(* IEC 61131-3 sources: Test-Git_ESME26/TestProgettoESME_26.fbsproj/AxisModuleLib Migration/AXM_FB_AxisModule.pou.xml.v3^ (part 2) *)

(* ---- Init_active.act.st ---- *)
__METADATA__
{
  "v3Meta": {
    "objectGuid": "f6f9ed11-c115-4c50-b3a9-4322940e64ce",
    "objectTypeGuid": "8ac092e5-3128-4e26-9e7e-11016c6684f2",
    "embeddedObjectTypeGuids": [
      "3b83b776-fb25-43b8-99f2-3c507c9143fc"
    ],
    "properties": {},
    "subObjects": {}
  }
}

iq_stStandardModuleItf.q_xActive := FALSE;
iq_stStandardModuleItf.q_xReady := FALSE;
iq_stStandardModuleItf.q_etDiag := GD.ET_Diag.Ok;
iq_stStandardModuleItf.q_udiDiagExt := AXM_ET_DiagExt.Disabled;
iq_stStandardModuleItf.q_sDiagExt := AXM_FC_EtDiagExtToString(i_etDiagExt := iq_stStandardModuleItf.q_udiDiagExt);
iq_stStandardModuleItf.q_sMsg := AXM_FC_EtDiagExtToString(i_etDiagExt := AXM_ET_DiagExt.Disabled);
iq_stStandardModuleItf.q_dwModuleType := TPL.ET_ModuleType.AxisModule;
iq_stStandardModuleItf.q_sModuleTypeName := 'AxisModule';
iq_stStandardModuleItf.q_udiModuleVersion := 1;

iq_stAxisModuleItf.stMain.q_etOpMode := AXM_ET_OpMode.NoOp;
iq_stAxisModuleItf.stMain.q_etState := AXM_ET_State.Disabled;

THIS^.DiagQuit();
THIS^.InactiveCMDExecution();

(* detect invalid configurations and avoid array index out of range error *)
IF(iq_stStandardModuleItf.iq_stExt.udiReactionOffset + TPL.ET_Reaction.MainsContactorOff > TPL.Gc_udiMaxNumberOfReactions) OR xExceptionReactionOutsideRange THEN (* module uses error reactions 1 to 5 *)
	xExceptionReactionOutsideRange := TRUE; (* create unquittable error *)
	(* create exception *)
	stExceptionInit.etDiag					:= GD.ET_Diag.InputParameterInvalid;
	stExceptionInit.udiDiagExt				:= AXM_ET_DiagExt.ReactionOffsetRange;
	stExceptionInit.sMsg					:= Standard.CONCAT('Value: ', UDINT_TO_STRING(iq_stStandardModuleItf.iq_stExt.udiReactionOffset));
	stExceptionInit.udiModuleId				:= iq_stStandardModuleItf.i_udiModuleId;
	stExceptionInit.sModuleName				:= iq_stStandardModuleItf.i_sModuleName;
	stExceptionInit.etSource				:= TPL.ET_ExceptionSource.AxisModule;
	stExceptionInit.timDelayTime			:= T#0MS;
	stExceptionInit.wHmiAttributes			:= 0;
	stExceptionInit.xAutoQuit				:= FALSE;
	stExceptionInit.stReaction.axReaction[TPL.ET_Reaction.AsyncStop]	:= TRUE; (* without offset on purpose *)
	iq_stStandardModuleItf.iq_stExt.udiReactionOffset := 0;
	ReportException(iq_stException := stExceptionInit);
ELSIF(iq_stStandardModuleItf.i_xEnable) THEN
	stReaction1 := stEmptyReaction;
	stReaction1.axReaction[iq_stStandardModuleItf.iq_stExt.udiReactionOffset + TPL.ET_Reaction.AsyncStop] := TRUE;
	stReaction2 := stEmptyReaction;
	stReaction2.axReaction[iq_stStandardModuleItf.iq_stExt.udiReactionOffset + TPL.ET_Reaction.SyncStopEL] := TRUE;
	stReaction3 := stEmptyReaction;
	stReaction3.axReaction[iq_stStandardModuleItf.iq_stExt.udiReactionOffset + TPL.ET_Reaction.SyncStopEH] := TRUE;
	stReaction4 := stEmptyReaction;
	stReaction4.axReaction[iq_stStandardModuleItf.iq_stExt.udiReactionOffset + TPL.ET_Reaction.StopEndOfCycle] := TRUE;

	(* Initialization of exception structures *)
	stExceptionCmdUnknown.etDiag			:= GD.ET_Diag.ExecutionAborted;
	stExceptionCmdUnknown.udiDiagExt		:= AXM_ET_DiagExt.CmdUnknown;
	stExceptionCmdUnknown.sMsg				:= 'Command unknown'; (* Replaced on usage *)
	stExceptionCmdUnknown.udiModuleId		:= iq_stStandardModuleItf.i_udiModuleId;
	stExceptionCmdUnknown.sModuleName		:= iq_stStandardModuleItf.i_sModuleName;
	stExceptionCmdUnknown.etSource			:= TPL.ET_ExceptionSource.AxisModule;
	stExceptionCmdUnknown.timDelayTime		:= T#0MS;
	stExceptionCmdUnknown.wHmiAttributes	:= 0;
	stExceptionCmdUnknown.xAutoQuit			:= FALSE;
	stExceptionCmdUnknown.stReaction		:= stReaction1;

	stExceptionCmdImpossibleOverwrite.etDiag			:= GD.ET_Diag.ExecutionAborted;
	stExceptionCmdImpossibleOverwrite.udiDiagExt		:= AXM_ET_DiagExt.CmdImpossibleOverwrite;
	stExceptionCmdImpossibleOverwrite.sMsg				:= 'Impossible command overwrite'; (* Replaced on usage *)
	stExceptionCmdImpossibleOverwrite.udiModuleId		:= iq_stStandardModuleItf.i_udiModuleId;
	stExceptionCmdImpossibleOverwrite.sModuleName		:= iq_stStandardModuleItf.i_sModuleName;
	stExceptionCmdImpossibleOverwrite.etSource			:= TPL.ET_ExceptionSource.AxisModule;
	stExceptionCmdImpossibleOverwrite.timDelayTime		:= T#0MS;
	stExceptionCmdImpossibleOverwrite.wHmiAttributes	:= 0;
	stExceptionCmdImpossibleOverwrite.xAutoQuit			:= FALSE;
	stExceptionCmdImpossibleOverwrite.stReaction		:= stReaction1;

	stExceptionCmdImpossibleState.etDiag			:= GD.ET_Diag.ExecutionAborted;
	stExceptionCmdImpossibleState.udiDiagExt		:= AXM_ET_DiagExt.CmdImpossibleState;
	stExceptionCmdImpossibleState.sMsg				:= 'Impossible command for state'; (* Replaced on usage *)
	stExceptionCmdImpossibleState.udiModuleId		:= iq_stStandardModuleItf.i_udiModuleId;
	stExceptionCmdImpossibleState.sModuleName		:= iq_stStandardModuleItf.i_sModuleName;
	stExceptionCmdImpossibleState.etSource			:= TPL.ET_ExceptionSource.AxisModule;
	stExceptionCmdImpossibleState.timDelayTime		:= T#0MS;
	stExceptionCmdImpossibleState.wHmiAttributes	:= 0;
	stExceptionCmdImpossibleState.xAutoQuit			:= FALSE;
	stExceptionCmdImpossibleState.stReaction		:= stReaction1;

	stWarningCmdImpossibleReaction.etDiag			:= GD.ET_Diag.ExecutionAborted;
	stWarningCmdImpossibleReaction.udiDiagExt		:= AXM_ET_DiagExt.CmdImpossibleReaction;
	stWarningCmdImpossibleReaction.sMsg				:= 'Impossible command on reaction'; (* Replaced on usage *)
	stWarningCmdImpossibleReaction.udiModuleId		:= iq_stStandardModuleItf.i_udiModuleId;
	stWarningCmdImpossibleReaction.sModuleName		:= iq_stStandardModuleItf.i_sModuleName;
	stWarningCmdImpossibleReaction.etSource			:= TPL.ET_ExceptionSource.AxisModule;
	stWarningCmdImpossibleReaction.timDelayTime	:= T#0MS;
	stWarningCmdImpossibleReaction.wHmiAttributes	:= 0;
	stWarningCmdImpossibleReaction.xAutoQuit		:= FALSE;

	stExceptionDriveFatal.etDiag			:= GD.ET_Diag.DriveConditionInvalid;
	stExceptionDriveFatal.udiDiagExt		:= AXM_ET_DiagExt.DriveExceptionFatal;
	stExceptionDriveFatal.sMsg				:= 'Drive diag'; (* Replaced on usage *)
	stExceptionDriveFatal.udiModuleId		:= iq_stStandardModuleItf.i_udiModuleId;
	stExceptionDriveFatal.sModuleName		:= iq_stStandardModuleItf.i_sModuleName;
	stExceptionDriveFatal.etSource			:= TPL.ET_ExceptionSource.AxisModule;
	stExceptionDriveFatal.timDelayTime		:= T#0MS;
	stExceptionDriveFatal.wHmiAttributes	:= 0;
	stExceptionDriveFatal.xAutoQuit			:= FALSE;
	stExceptionDriveFatal.stReaction		:= stReaction1;

	stExcepitonDrive.etDiag			:= GD.ET_Diag.DriveConditionInvalid;
	stExcepitonDrive.udiDiagExt		:= AXM_ET_DiagExt.DriveException;
	stExcepitonDrive.sMsg			:= 'Drive diag'; (* Replaced on usage *)
	stExcepitonDrive.udiModuleId	:= iq_stStandardModuleItf.i_udiModuleId;
	stExcepitonDrive.sModuleName	:= iq_stStandardModuleItf.i_sModuleName;
	stExcepitonDrive.etSource		:= TPL.ET_ExceptionSource.AxisModule;
	stExcepitonDrive.timDelayTime	:= T#0MS;
	stExcepitonDrive.wHmiAttributes	:= 0;
	stExcepitonDrive.xAutoQuit		:= FALSE;
	stExcepitonDrive.stReaction		:= stReaction2;

	stWarningDrive.etDiag			:= GD.ET_Diag.DriveConditionInvalid;
	stWarningDrive.udiDiagExt		:= AXM_ET_DiagExt.DriveWarning;
	stWarningDrive.sMsg				:= 'Drive warning'; (* Replaced on usage *)
	stWarningDrive.udiModuleId		:= iq_stStandardModuleItf.i_udiModuleId;
	stWarningDrive.sModuleName		:= iq_stStandardModuleItf.i_sModuleName;
	stWarningDrive.etSource			:= TPL.ET_ExceptionSource.AxisModule;
	stWarningDrive.timDelayTime		:= T#0MS;
	stWarningDrive.wHmiAttributes	:= 0;
	stWarningDrive.xAutoQuit		:= FALSE;
	stWarningDrive.stReaction		:= stReaction4;

	stExceptionPosHwLimit.etDiag			:= GD.ET_Diag.LimitReached;
	stExceptionPosHwLimit.udiDiagExt		:= AXM_ET_DiagExt.HwLimitPosReached;
	stExceptionPosHwLimit.sMsg				:= '';
	stExceptionPosHwLimit.udiModuleId		:= iq_stStandardModuleItf.i_udiModuleId;
	stExceptionPosHwLimit.sModuleName		:= iq_stStandardModuleItf.i_sModuleName;
	stExceptionPosHwLimit.etSource			:= TPL.ET_ExceptionSource.AxisModule;
	stExceptionPosHwLimit.timDelayTime		:= T#0MS;
	stExceptionPosHwLimit.wHmiAttributes	:= 0;
	stExceptionPosHwLimit.xAutoQuit			:= FALSE;
	stExceptionPosHwLimit.stReaction		:= stReaction3;

	stExceptionNegHwLimit.etDiag			:= GD.ET_Diag.LimitReached;
	stExceptionNegHwLimit.udiDiagExt		:= AXM_ET_DiagExt.HwLimitNegReached;
	stExceptionNegHwLimit.sMsg				:= '';
	stExceptionNegHwLimit.udiModuleId		:= iq_stStandardModuleItf.i_udiModuleId;
	stExceptionNegHwLimit.sModuleName		:= iq_stStandardModuleItf.i_sModuleName;
	stExceptionNegHwLimit.etSource			:= TPL.ET_ExceptionSource.AxisModule;
	stExceptionNegHwLimit.timDelayTime		:= T#0MS;
	stExceptionNegHwLimit.wHmiAttributes	:= 0;
	stExceptionNegHwLimit.xAutoQuit			:= FALSE;
	stExceptionNegHwLimit.stReaction		:= stReaction3;

	stWarningPosHwLimit.etDiag			:= GD.ET_Diag.LimitReached;
	stWarningPosHwLimit.udiDiagExt		:= AXM_ET_DiagExt.HwLimitPosWarning;
	stWarningPosHwLimit.sMsg			:= '';
	stWarningPosHwLimit.udiModuleId		:= iq_stStandardModuleItf.i_udiModuleId;
	stWarningPosHwLimit.sModuleName		:= iq_stStandardModuleItf.i_sModuleName;
	stWarningPosHwLimit.etSource		:= TPL.ET_ExceptionSource.AxisModule;
	stWarningPosHwLimit.timDelayTime	:= T#0MS;
	stWarningPosHwLimit.wHmiAttributes	:= 0;
	stWarningPosHwLimit.xAutoQuit		:= TRUE;

	stWarningNegHwLimit.etDiag			:= GD.ET_Diag.LimitReached;
	stWarningNegHwLimit.udiDiagExt		:= AXM_ET_DiagExt.HwLimitNegWarning;
	stWarningNegHwLimit.sMsg			:= '';
	stWarningNegHwLimit.udiModuleId		:= iq_stStandardModuleItf.i_udiModuleId;
	stWarningNegHwLimit.sModuleName		:= iq_stStandardModuleItf.i_sModuleName;
	stWarningNegHwLimit.etSource		:= TPL.ET_ExceptionSource.AxisModule;
	stWarningNegHwLimit.timDelayTime	:= T#0MS;
	stWarningNegHwLimit.wHmiAttributes	:= 0;
	stWarningNegHwLimit.xAutoQuit		:= TRUE;

	stExceptionVelLimitCrossed.etDiag			:= GD.ET_Diag.LimitReached;
	stExceptionVelLimitCrossed.udiDiagExt		:= AXM_ET_DiagExt.ReducedVelocityLImit;
	stExceptionVelLimitCrossed.sMsg				:= '';
	stExceptionVelLimitCrossed.udiModuleId		:= iq_stStandardModuleItf.i_udiModuleId;
	stExceptionVelLimitCrossed.sModuleName		:= iq_stStandardModuleItf.i_sModuleName;
	stExceptionVelLimitCrossed.etSource			:= TPL.ET_ExceptionSource.AxisModule;
	stExceptionVelLimitCrossed.timDelayTime		:= T#0MS;
	stExceptionVelLimitCrossed.wHmiAttributes	:= 0;
	stExceptionVelLimitCrossed.xAutoQuit		:= FALSE;
	stExceptionVelLimitCrossed.stReaction		:= stReaction1;

	stExceptionUnexpected.etDiag			:= GD.ET_Diag.UnexpectedProgramBehavior;
	stExceptionUnexpected.udiDiagExt		:= AXM_ET_DiagExt.UnknownFeedback;
	stExceptionUnexpected.sMsg				:= ''; (* Replaced on usage *)
	stExceptionUnexpected.udiModuleId		:= iq_stStandardModuleItf.i_udiModuleId;
	stExceptionUnexpected.sModuleName		:= iq_stStandardModuleItf.i_sModuleName;
	stExceptionUnexpected.etSource			:= TPL.ET_ExceptionSource.AxisModule;
	stExceptionUnexpected.timDelayTime		:= T#0MS;
	stExceptionUnexpected.wHmiAttributes	:= 0;
	stExceptionUnexpected.xAutoQuit			:= FALSE;
	stExceptionUnexpected.stReaction		:= stReaction1;

	stExceptionModuleReaction1.etDiag			:= GD.ET_Diag.InputParameterInvalid;(* Replaced on usage *)
	stExceptionModuleReaction1.udiDiagExt		:= AXM_ET_DiagExt.DriveInvalid;(* Replaced on usage *)
	stExceptionModuleReaction1.sMsg				:= '';(* Replaced on usage *)
	stExceptionModuleReaction1.udiModuleId		:= iq_stStandardModuleItf.i_udiModuleId;
	stExceptionModuleReaction1.sModuleName		:= iq_stStandardModuleItf.i_sModuleName;
	stExceptionModuleReaction1.etSource			:= TPL.ET_ExceptionSource.AxisModule;
	stExceptionModuleReaction1.timDelayTime		:= T#0MS;
	stExceptionModuleReaction1.wHmiAttributes	:= 0;
	stExceptionModuleReaction1.xAutoQuit		:= FALSE;
	stExceptionModuleReaction1.stReaction		:= stReaction1;

	stExceptionModuleReaction2.etDiag			:= GD.ET_Diag.InputParameterInvalid;(* Replaced on usage *)
	stExceptionModuleReaction2.udiDiagExt		:= AXM_ET_DiagExt.DriveInvalid;(* Replaced on usage *)
	stExceptionModuleReaction2.sMsg				:= '';(* Replaced on usage *)
	stExceptionModuleReaction2.udiModuleId		:= iq_stStandardModuleItf.i_udiModuleId;
	stExceptionModuleReaction2.sModuleName		:= iq_stStandardModuleItf.i_sModuleName;
	stExceptionModuleReaction2.etSource			:= TPL.ET_ExceptionSource.AxisModule;
	stExceptionModuleReaction2.timDelayTime		:= T#0MS;
	stExceptionModuleReaction2.wHmiAttributes	:= 0;
	stExceptionModuleReaction2.xAutoQuit		:= FALSE;
	stExceptionModuleReaction2.stReaction		:= stReaction2;

	stExceptionModuleReaction3.etDiag			:= GD.ET_Diag.InputParameterInvalid;(* Replaced on usage *)
	stExceptionModuleReaction3.udiDiagExt		:= AXM_ET_DiagExt.DriveInvalid;(* Replaced on usage *)
	stExceptionModuleReaction3.sMsg				:= '';(* Replaced on usage *)
	stExceptionModuleReaction3.udiModuleId		:= iq_stStandardModuleItf.i_udiModuleId;
	stExceptionModuleReaction3.sModuleName		:= iq_stStandardModuleItf.i_sModuleName;
	stExceptionModuleReaction3.etSource			:= TPL.ET_ExceptionSource.AxisModule;
	stExceptionModuleReaction3.timDelayTime		:= T#0MS;
	stExceptionModuleReaction3.wHmiAttributes	:= 0;
	stExceptionModuleReaction3.xAutoQuit		:= FALSE;
	stExceptionModuleReaction3.stReaction		:= stReaction3;

	stExceptionModuleReaction4.etDiag			:= GD.ET_Diag.InputParameterInvalid;(* Replaced on usage *)
	stExceptionModuleReaction4.udiDiagExt		:= AXM_ET_DiagExt.DriveInvalid;(* Replaced on usage *)
	stExceptionModuleReaction4.sMsg				:= '';(* Replaced on usage *)
	stExceptionModuleReaction4.udiModuleId		:= iq_stStandardModuleItf.i_udiModuleId;
	stExceptionModuleReaction4.sModuleName		:= iq_stStandardModuleItf.i_sModuleName;
	stExceptionModuleReaction4.etSource			:= TPL.ET_ExceptionSource.AxisModule;
	stExceptionModuleReaction4.timDelayTime		:= T#0MS;
	stExceptionModuleReaction4.wHmiAttributes	:= 0;
	stExceptionModuleReaction4.xAutoQuit		:= FALSE;
	stExceptionModuleReaction4.stReaction		:= stReaction4;

	IF (iq_stAxisModuleItf.stMain.i_ifDrive = 0) THEN
		stExceptionModuleReaction1.etDiag		:= GD.ET_Diag.InputParameterInvalid;
		stExceptionModuleReaction1.udiDiagExt	:= AXM_ET_DiagExt.DriveInvalid;
		stExceptionModuleReaction1.sMsg			:= 'No drive given';
		ReportException(iq_stException := stExceptionModuleReaction1);
	ELSE
		iq_stStandardModuleItf.q_xActive := TRUE;
		FOR udii := 1 TO TPL.Gc_udiMaxNumberOfReactions DO
			stLocalReaction.axReaction[udii] := FALSE;
		END_FOR
		xSuccess := __QUERYINTERFACE(iq_stAxisModuleItf.stMain.i_ifDrive, ifGetParentDevice);
		IF xSuccess THEN
			ifDeviceAccess := ifGetParentDevice.GetParentDevice();
			xSuccess := __QUERYINTERFACE(ifDeviceAccess, ifDeviceTreeObjectAccess);
			IF xSuccess THEN
				iq_stAxisModuleItf.stMain.q_sDriveName := ifDeviceTreeObjectAccess.DeviceTreeObject.Name;
			END_IF
		ELSE
			//no device tree object
			iq_stAxisModuleItf.stMain.q_sDriveName := '';
		END_IF
		xEnableFlag := TRUE;

		stCamTab:=	iq_stAxisModuleItf.stMultiCam.iq_astMotionPar[AXM_ET_ParId.Idle];
		xInitHomingDone := FALSE;
		udiInitHoming := 0;
		iq_stAxisModuleItf.stMain.q_etState := AXM_ET_State.Initializing;
		xStartBitLastCycle := FALSE;
		etPowerState := AXM_ET_PowerState.PowerOff;

		IF fbLoggerPoint.etLogLevel >= APL.ET_LogLevel.UserAction THEN
			fbLoggerPoint.AddLogEntry(	i_etLogLevel	:= APL.ET_LogLevel.UserAction,
										i_etDiag		:= GD.ET_Diag.Ok,
										i_udiDiagExt	:= AXM_ET_DiagExt.Ok,
										i_sMessage		:= 'enabeling Module',
										q_etDiag		:= ,
										q_etDiagExt		:= );
		END_IF
		fbDriveEnable.RegisterLoggerPoint(	i_ifParent	:= fbLoggerPoint,
											i_sName		:= 'DriveEnable',
											q_etDiag	=> ,
											q_etDiagExt => );
	END_IF

END_IF
THIS^.Output_active();

(* ---- InitHoming_active.act.st ---- *)
__METADATA__
{
  "v3Meta": {
    "objectGuid": "dae82e5a-5072-46fa-9bd0-11e67c638b29",
    "objectTypeGuid": "8ac092e5-3128-4e26-9e7e-11016c6684f2",
    "embeddedObjectTypeGuids": [
      "3b83b776-fb25-43b8-99f2-3c507c9143fc"
    ],
    "properties": {},
    "subObjects": {}
  }
}

InactiveCMDExecution();

fbHome.stReducedVelocity := iq_stAxisModuleItf.stMain.stReducedVelocity;
IF iq_stAxisModuleItf.stHome.i_etMode = PDL_ET_HomeMode.RestorePosFromAxisEncoder
	OR iq_stAxisModuleItf.stHome.i_etMode = PDL_ET_HomeMode.WriteAxisEncoder THEN
	etHomeModeTemp := PDL_ET_HomeMode.RestorePosFromAxisEncoder;
ELSE
	etHomeModeTemp := PDL_ET_HomeMode.RestorePosFromRetain;
END_IF
IF iq_stAxisModuleItf.stHome.i_xEnableInitAbsReadPos AND ( (etHomeModeTemp = PDL_ET_HomeMode.RestorePosFromAxisEncoder) OR
															(etHomeModeTemp = PDL_ET_HomeMode.RestorePosFromRetain) ) THEN
	stFbHomeSetPosProperty.i_lrAbsEncOffset			:= iq_stAxisModuleItf.stHome.stSetPos.i_lrAbsEncOffset;
	stFbHomeSetPosProperty.i_lrEncoderPosition		:= iq_stAxisModuleItf.stHome.stSetPos.i_lrEncoderPosition;
	stFbHomeSetPosProperty.i_lrHomePosition			:= iq_stAxisModuleItf.stHome.stSetPos.i_lrHomePosition;
	stFbHomeSetPosProperty.i_lrRestoreWindow		:= iq_stAxisModuleItf.stHome.stSetPos.i_lrRestoreWindow;
	stFbHomeSetPosProperty.i_lrUserPeriod			:= iq_stAxisModuleItf.stHome.stSetPos.i_lrUserPeriod;
	stFbHomeSetPosProperty.iq_pstRestorePosRetain	:= iq_stAxisModuleItf.stHome.stSetPos.iq_pstRestorePosRetain;
	stFbHomeSetPosProperty.iq_lencAxis				:= iq_stAxisModuleItf.stMain.iq_lencEncoder;
	fbHome.stSetPos := stFbHomeSetPosProperty;

	IF NOT iq_stAxisModuleItf.stHome.stSetPos.i_xKeepPowerDisabled AND
			udiInitHoming = 0 AND
			iq_stAxisModuleItf.stMain.i_ifDrive.etAxisState >= MOIN.ET_AxisState.Standstill THEN
		//Create LoggerEnty
		ReadTrackingDeviation(q_sLrealConversion => sLrealConversion);

		fbLoggerPoint.AddLogEntry (
				i_etLogLevel 	:= APL.ET_LogLevel.StatusMessage,
				i_etDiag		:= GD.ET_Diag.Ok,
				i_udiDiagExt	:= 0,
				i_sMessage		:= Standard.CONCAT('SetPos-Homing in Init:  Axis-State >= Standstill; TrackingDeviation: ',sLrealConversion)
			);
			udiInitHoming := 30;
	ELSIF udiInitHoming = 0 THEN
		IF 	iq_stAxisModuleItf.stMain.i_ifDrive.etAxisState >= MOIN.ET_AxisState.Standstill THEN
			udiInitHoming := 10;
		ELSE
			udiInitHoming := 30;
		END_IF
	END_IF

	CASE udiInitHoming OF
	0:
		udiInitHoming := 30;
		;
	10: (* Disable Power if i_xKeepPowerDisabled is set*)
		IF iq_stAxisModuleItf.stHome.stSetPos.i_xKeepPowerDisabled THEN
			fbDriveEnable(	i_xEnable		:= TRUE,
							i_ifDrive		:= iq_stAxisModuleItf.stMain.i_ifDrive,
							i_xEnableDrive	:= FALSE,
							i_xDiagQuit		:= iq_stStandardModuleItf.i_xDiagQuit,
							q_xActive		=> ,
							q_xReady		=> ,
							q_etDiag		=> etDiagBuffer,
							q_etDiagExt		=> etDiagExtBufferPDL,
							q_sMsg			=> sDiagMsgBuffer,
							q_xDriveEnabled	=> );
			IF (etDiagBuffer <> GD.ET_Diag.Ok) THEN
				DiagTestDriveEnable(	iq_etDiag		:= fbDriveEnable.q_etDiag,
										iq_etDiagExt	:= fbDriveEnable.q_etDiagExt,
										iq_sMsg			:= fbDriveEnable.q_sMsg);
				udiInitHoming := 30;
			END_IF

			IF fbDriveEnable.q_xActive AND NOT fbDriveEnable.q_xDriveEnabled THEN
				fbDriveEnable(	i_xEnable		:= FALSE);
				udiInitHoming := 20;
			END_IF
		ELSE
			udiInitHoming := 30;
		END_IF

	20: (* Check FB_DriveEnable disabled *)
		IF NOT fbDriveEnable.q_xActive THEN
			udiInitHoming := 30;
		END_IF

	30: (* Do initial homing *)
		fbHome(	i_xEnable				:= TRUE,
				i_etMode				:= etHomeModeTemp,
				i_ifDrive	 			:= iq_stAxisModuleItf.stMain.i_ifDrive,
				i_xHwLimitNeg			:= FALSE,
				i_xHwLimitPos			:= FALSE,
				i_xStart				:= TRUE,
				q_xActive				=> ,
				q_xReady				=> ,
				q_etDiag				=> etDiagBuffer,
				q_etDiagExt				=> etDiagExtBufferPDL,
				q_sMsg					=> sDiagMsgBuffer,
				q_xDisableDrive			=> ,
				q_xMotionInstructionActive	=> ,
				q_lrPosition			=> ,
				q_lrEncoderPosition		=> ,
				q_xHomeOk				=> );
		IF (fbHome.q_etDiag <> GD.ET_Diag.Ok) THEN
			DiagTestHoming(	iq_etDiag		:= fbHome.q_etDiag,
							iq_etDiagExt	:= fbHome.q_etDiagExt,
							iq_sMsg			:= fbHome.q_sMsg);
			udiInitHoming := 40;
		END_IF

		IF fbHome.q_xHomeOk THEN
			iq_stAxisModuleItf.stMain.q_xHomeOk := TRUE;
			IF fbLoggerPoint.etLogLevel >= APL.ET_LogLevel.StatusMessage THEN
				IF (etHomeModeTemp = PDL_ET_HomeMode.RestorePosFromAxisEncoder) THEN
					fbLoggerPoint.AddLogEntry(	i_etLogLevel	:= APL.ET_LogLevel.StatusMessage,
												i_etDiag		:= GD.ET_Diag.Ok,
												i_udiDiagExt	:= AXM_ET_DiagExt.Ok,
												i_sMessage		:= 'InitAbsReadPos done from AxisEncoder',
												q_etDiag		:= ,
												q_etDiagExt		:= );
				ELSE
					fbLoggerPoint.AddLogEntry(	i_etLogLevel	:= APL.ET_LogLevel.StatusMessage,
												i_etDiag		:= GD.ET_Diag.Ok,
												i_udiDiagExt	:= AXM_ET_DiagExt.Ok,
												i_sMessage		:= 'InitAbsReadPos done from Retain',
												q_etDiag		:= ,
												q_etDiagExt		:= );
				END_IF
			END_IF
			udiInitHoming := 40;
		END_IF

	40: (* clean up initial Homing *)
		fbHome(	i_xEnable				:= FALSE,
				i_etMode				:= etHomeModeTemp,
				i_ifDrive	 			:= iq_stAxisModuleItf.stMain.i_ifDrive,
				i_xHwLimitNeg			:= FALSE,
				i_xHwLimitPos			:= FALSE,
				i_xStart				:= FALSE,
				q_xActive				=> ,
				q_xReady				=> ,
				q_etDiag				=> etDiagBuffer,
				q_etDiagExt				=> etDiagExtBufferPDL,
				q_sMsg					=> sDiagMsgBuffer,
				q_xDisableDrive			=> ,
				q_xMotionInstructionActive	=> ,
				q_lrPosition			=> ,
				q_lrEncoderPosition		=> ,
				q_xHomeOk				=> );
		IF (fbHome.q_etDiag <> GD.ET_Diag.Ok) THEN
			DiagTestHoming(	iq_etDiag		:= fbHome.q_etDiag,
							iq_etDiagExt	:= fbHome.q_etDiagExt,
							iq_sMsg			:= fbHome.q_sMsg);
			xInitHomingDone := TRUE;
		END_IF
		IF NOT fbHome.q_xActive THEN
			xInitHomingDone := TRUE;
		END_IF

	END_CASE

ELSE
	xInitHomingDone := TRUE;
END_IF
THIS^.Output_active();

(* ---- Input_active.act.st ---- *)
__METADATA__
{
  "v3Meta": {
    "objectGuid": "61561b81-6e46-47b7-b302-ee9f18f8c31f",
    "objectTypeGuid": "8ac092e5-3128-4e26-9e7e-11016c6684f2",
    "embeddedObjectTypeGuids": [
      "3b83b776-fb25-43b8-99f2-3c507c9143fc"
    ],
    "properties": {},
    "subObjects": {}
  }
}

IF iq_stAxisModuleItf.stHome.i_xResetHomeOk THEN
	iq_stAxisModuleItf.stMain.q_xHomeOk := FALSE;

	IF fbHome.q_xHomeOk = TRUE THEN
		xResetHomeOkActive := TRUE;
	END_IF
END_IF

(* -----------------------------------------------------------------------------------------------*)
(* Check DiagQuit *)
(* -----------------------------------------------------------------------------------------------*)
THIS^.DiagQuit();

(* -----------------------------------------------------------------------------------------------*)
(* Check external Reaction *)
(* -----------------------------------------------------------------------------------------------*)

stModuleReaction.axReaction[TPL.ET_Reaction.AsyncStop] := stLocalReaction.axReaction[TPL.ET_Reaction.AsyncStop] OR iq_stStandardModuleItf.i_stReaction.axReaction[TPL.ET_Reaction.AsyncStop];
stModuleReaction.axReaction[TPL.ET_Reaction.SyncStopEL] := stLocalReaction.axReaction[TPL.ET_Reaction.SyncStopEL] OR iq_stStandardModuleItf.i_stReaction.axReaction[TPL.ET_Reaction.SyncStopEL];
stModuleReaction.axReaction[TPL.ET_Reaction.SyncStopEH] := stLocalReaction.axReaction[TPL.ET_Reaction.SyncStopEH] OR iq_stStandardModuleItf.i_stReaction.axReaction[TPL.ET_Reaction.SyncStopEH];
stModuleReaction.axReaction[TPL.ET_Reaction.StopEndOfCycle] := stLocalReaction.axReaction[TPL.ET_Reaction.StopEndOfCycle] OR iq_stStandardModuleItf.i_stReaction.axReaction[TPL.ET_Reaction.StopEndOfCycle];
stModuleReaction.axReaction[TPL.ET_Reaction.MainsContactorOff] := stLocalReaction.axReaction[TPL.ET_Reaction.MainsContactorOff] OR iq_stStandardModuleItf.i_stReaction.axReaction[TPL.ET_Reaction.MainsContactorOff];

(* -----------------------------------------------------------------------------------------------*)
(* save axis pos in case of restore position *)
(* -----------------------------------------------------------------------------------------------*)
IF (iq_stAxisModuleItf.stMain.i_ifDrive = 0) THEN
	stExceptionModuleReaction1.etDiag		:= GD.ET_Diag.InputParameterInvalid;
	stExceptionModuleReaction1.udiDiagExt	:= AXM_ET_DiagExt.DriveInvalid;
	stExceptionModuleReaction1.sMsg			:= 'No drive given';
	ReportException(iq_stException := stExceptionModuleReaction1);

	etPowerState					:= AXM_ET_PowerState.PowerOff;
	xCMDPowerOn						:= FALSE;

(*** save axis pos in case of restore position ***)
ELSIF iq_stAxisModuleItf.stHome.i_xEnableInitAbsReadPos AND
	iq_stAxisModuleItf.stHome.i_etMode <> PDL_ET_HomeMode.RestorePosFromAxisencoder AND
	iq_stAxisModuleItf.stHome.i_etMode <> PDL_ET_HomeMode.WriteAxisEncoder AND
	iq_stAxisModuleItf.stMain.q_xHomeOk THEN

	IF (iq_stAxisModuleItf.stHome.stSetPos.iq_pstRestorePosRetain <= 0) THEN
		stExceptionModuleReaction3.etDiag := GD.ET_Diag.InputParameterInvalid;
		stExceptionModuleReaction3.udiDiagExt := PDL_ET_DiagExt.PointerRestorePosRetainInvalid;
		stExceptionModuleReaction3.sMsg := 'pointer is zero';
		ReportException(iq_stException := stExceptionModuleReaction3);

		etPowerState					:= AXM_ET_PowerState.PowerOff;
		xCMDPowerOn						:= FALSE;
	ELSIF (FC_GetSercosState() = SMI.ET_SercosState.Phase4) THEN
		PDL_FC_SaveAxisPosition(	i_etPosType				:= PDL_ET_PosType.MechPosition,
									i_ifDrive				:= iq_stAxisModuleItf.stMain.i_ifDrive,
									iq_stRestorePosition	:= iq_stAxisModuleItf.stHome.stSetPos.iq_pstRestorePosRetain^,
									q_etDiag				=> etDiagBuffer,
									q_etDiagExt				=> etDiagExtBufferPDL,
									q_sMsg					=> sDiagMsgBuffer);
		IF (etDiagBuffer <> GD.ET_Diag.Ok) THEN
			stExceptionUnexpected.udiDiagExt := AXM_ET_DiagExt.UnexpectedFeedback;
			stExceptionUnexpected.sMsg := SE_CTBX.FC_MultiConcat(	i_sString1 := 'FC_SaveAxisPosition ',
																i_sString2 := PDL_FC_EtDiagExtToString(i_etDiagExt := etDiagExtBufferPDL),
																i_sString3 := ' ',
																i_sString4 := sDiagMsgBuffer);
			ReportException(iq_stException := stExceptionUnexpected);
		END_IF
	END_IF
END_IF

(* ---- Logging_active.act.st ---- *)
__METADATA__
{
  "v3Meta": {
    "objectGuid": "20ce76ab-1f0b-407f-9e41-8519cd1cefc9",
    "objectTypeGuid": "8ac092e5-3128-4e26-9e7e-11016c6684f2",
    "embeddedObjectTypeGuids": [
      "3b83b776-fb25-43b8-99f2-3c507c9143fc"
    ],
    "properties": {},
    "subObjects": {}
  }
}

(* System generated code, do not change without consulting Schneider Electric - otherwise you risk instability!!!*)

fbLogger(		i_xEnable			:= iq_stStandardModuleItf.i_xLogEnable,
				i_wLogDataFilter	:= iq_stStandardModuleItf.i_wLogDataFilter,
				i_sModuleName		:= iq_stStandardModuleItf.i_sModuleName,
				i_udiModuleId		:= iq_stStandardModuleItf.i_udiModuleId,
				i_diCmd				:= iq_stStandardModuleItf.iq_diCmd,
				i_diStartStep		:= 0,
				i_stReaction		:= iq_stStandardModuleItf.i_stReaction,
				iq_stExceptionList	:= iq_stExceptionList,
				iq_stLogDataList	:= iq_stLogDataList,
				q_xActive			=> xLogger_Active,
				q_xReady			=> ,
				q_etDiag			=> ,
				q_etDiagExt			=> );

IF iq_stAxisModuleItf.stMain.stReducedVelocity.i_xEnableReducedVelocity AND NOT xReducedEnableFlag THEN
	xReducedEnableFlag:=TRUE;
	xOnlyLimitCheckFlag:=NOT iq_stAxisModuleItf.stMain.stReducedVelocity.i_xOnlyLimitCheck;
ELSIF NOT iq_stAxisModuleItf.stMain.stReducedVelocity.i_xEnableReducedVelocity AND  xReducedEnableFlag THEN
	xReducedEnableFlag:=FALSE;
		TPL.FC_GetTimeStamp(	q_etDiag	=> ,
								q_etDiagExt	=> ,
								q_sMsg		=> ,
								q_dateDate	=> dateNow,
								q_todTime	=> todNow);
		TPL.FC_SingleLoggerEntry(		i_etReason		:= TPL.ET_LogDataFilter.User,
										i_dateDate		:= dateNow,
										i_todTime		:= todNow,
										i_udiModuleId	:= iq_stStandardModuleItf.i_udiModuleId,
										i_sModuleName	:= iq_stStandardModuleItf.i_sModuleName,
										i_diCmd			:= 0,
										i_diStartStep	:= 0,
										i_stReaction	:= stEmptyReaction,
										i_etDiag		:= 0,
										i_udiDiagExt	:= 0,
										i_sDiagExt		:= '',
										i_sMsg			:= 'Reduced Velocity Off',
										i_etSource		:= TPL.ET_ExceptionSource.AxisModule,
										i_xAutoQuit		:= FALSE,
										iq_stLogDataList:= iq_stLogDataList,
										q_etDiag		=> ,
										q_etDiagExt		=> );
END_IF

IF xReducedEnableFlag THEN
	IF iq_stAxisModuleItf.stMain.stReducedVelocity.i_xOnlyLimitCheck  AND NOT xOnlyLimitCheckFlag THEN
		xOnlyLimitCheckFlag:=TRUE;
		TPL.FC_GetTimeStamp(	q_etDiag	=> ,
								q_etDiagExt	=> ,
								q_sMsg		=> ,
								q_dateDate	=> dateNow,
								q_todTime	=> todNow);
		TPL.FC_SingleLoggerEntry(		i_etReason		:= TPL.ET_LogDataFilter.User,
										i_dateDate		:= dateNow,
										i_todTime		:= todNow,
										i_udiModuleId	:= iq_stStandardModuleItf.i_udiModuleId,
										i_sModuleName	:= iq_stStandardModuleItf.i_sModuleName,
										i_diCmd			:= 0,
										i_diStartStep	:= 0,
										i_stReaction	:= stEmptyReaction,
										i_etDiag		:= 0,
										i_udiDiagExt	:= 0,
										i_sDiagExt		:= '',
										i_sMsg			:= 'Reduced Velocity On; only Limit check',
										i_etSource		:= TPL.ET_ExceptionSource.AxisModule,
										i_xAutoQuit		:= FALSE,
										iq_stLogDataList:= iq_stLogDataList,
										q_etDiag		=> ,
										q_etDiagExt		=> );
	ELSIF NOT iq_stAxisModuleItf.stMain.stReducedVelocity.i_xOnlyLimitCheck  AND  xOnlyLimitCheckFlag THEN
		xOnlyLimitCheckFlag:=FALSE;
		TPL.FC_GetTimeStamp(	q_etDiag	=> ,
								q_etDiagExt	=> ,
								q_sMsg		=> ,
								q_dateDate	=> dateNow,
								q_todTime	=> todNow);
		TPL.FC_SingleLoggerEntry(		i_etReason		:= TPL.ET_LogDataFilter.User,
										i_dateDate		:= dateNow,
										i_todTime		:= todNow,
										i_udiModuleId	:= iq_stStandardModuleItf.i_udiModuleId,
										i_sModuleName	:= iq_stStandardModuleItf.i_sModuleName,
										i_diCmd			:= 0,
										i_diStartStep	:= 0,
										i_stReaction	:= stEmptyReaction,
										i_etDiag		:= 0,
										i_udiDiagExt	:= 0,
										i_sDiagExt		:= '',
										i_sMsg			:= 'Reduced Velocity On; with limitation',
										i_etSource		:= TPL.ET_ExceptionSource.AxisModule,
										i_xAutoQuit		:= FALSE,
										iq_stLogDataList:= iq_stLogDataList,
										q_etDiag		=> ,
										q_etDiagExt		=> );
	END_IF
END_IF

(* End of system generated code, do not change without consulting Schneider Electric - otherwise you risk instability!!!*)

(* ---- Manual_active.act.st ---- *)
__METADATA__
{
  "v3Meta": {
    "objectGuid": "e5dd1cdc-5ee5-46d9-a02c-cd1dfda45dfe",
    "objectTypeGuid": "8ac092e5-3128-4e26-9e7e-11016c6684f2",
    "embeddedObjectTypeGuids": [
      "3b83b776-fb25-43b8-99f2-3c507c9143fc"
    ],
    "properties": {},
    "subObjects": {}
  }
}

iq_stAxisModuleItf.stMain.q_etOpMode := AXM_ET_OpMode.Manual;

xManJogForw :=
	(iq_stAxisModuleItf.stManual.i_xJogForw AND
		NOT iq_stAxisModuleItf.stMain.i_xHwLimitPos AND
		NOT stModuleReaction.axReaction[TPL.ET_Reaction.StopEndOfCycle]);
xManJogBack :=
	(iq_stAxisModuleItf.stManual.i_xJogBack AND
		NOT iq_stAxisModuleItf.stMain.i_xHwLimitNeg AND
		NOT stModuleReaction.axReaction[TPL.ET_Reaction.StopEndOfCycle]);

IF (iq_stAxisModuleItf.stMain.stReducedVelocity.i_xEnableReducedVelocity AND NOT iq_stAxisModuleItf.stMain.stReducedVelocity.i_xOnlyLimitCheck) THEN

	lrManVel := MIN(iq_stAxisModuleItf.stManual.i_lrVel, iq_stAxisModuleItf.stMain.stReducedVelocity.i_lrMaxReducedVelocity);
ELSE
	lrManVel := iq_stAxisModuleItf.stManual.i_lrVel;
END_IF

fbJogging(
	i_xEnable                  := xManEnable AND fbDriveEnable.q_xDriveEnabled,
	i_ifDrive                  := iq_stAxisModuleItf.stMain.i_ifDrive,
	i_xJogForw                 := xManJogForw,
	i_xJogBack                 := xManJogBack,
	i_lrPeriod                 := iq_stAxisModuleItf.stManual.i_lrPeriod,
	i_xEndless                 := iq_stAxisModuleItf.stManual.i_xEndless,
	i_lrMaxDistance            := iq_stAxisModuleItf.stManual.i_lrMaxDistance,
	i_lrVel                    := lrManVel,
	i_lrAcc                    := iq_stAxisModuleItf.stManual.i_lrAcc,
	i_lrDec                    := iq_stAxisModuleItf.stManual.i_lrDec,
	i_lrJerk                   := iq_stAxisModuleItf.stManual.i_lrJerk,
	q_xActive                  =>,
	q_xReady                   =>,
	q_etDiag                   => etDiagBuffer,
	q_etDiagExt                => etDiagExtBufferPDL,
	q_sMsg                     => sDiagMsgBuffer,
	q_xMotionInstructionActive =>,
	q_lrPosition               =>,
	q_xStepFinished            =>
);

DiagTestJogging(iq_etDiag := fbJogging.q_etDiag, iq_etDiagExt := fbJogging.q_etDiagExt, iq_sMsg := fbJogging.q_sMsg);

IF fbJogging.q_xReady THEN
	iq_stAxisModuleItf.stMain.q_etState := AXM_ET_State.ManualRunning;
ELSE
	IF xManEnable THEN
		iq_stAxisModuleItf.stMain.q_etState := AXM_ET_State.ManualInit;
	ELSE
		iq_stAxisModuleItf.stMain.q_etState := AXM_ET_State.ManualExit;
	END_IF
END_IF

IF NOT xManEnable AND NOT fbJogging.q_xActive THEN
	xManActive := FALSE;
END_IF

(* ---- MultiCam_active.act.st ---- *)
__METADATA__
{
  "v3Meta": {
    "objectGuid": "5e85057d-b7e3-4f89-8b75-5d4e0717c30c",
    "objectTypeGuid": "8ac092e5-3128-4e26-9e7e-11016c6684f2",
    "embeddedObjectTypeGuids": [
      "3b83b776-fb25-43b8-99f2-3c507c9143fc"
    ],
    "properties": {},
    "subObjects": {}
  }
}

iq_stAxisModuleItf.stMain.q_etOpMode := AXM_ET_OpMode.MultiCam;

xEnableMultiCamFb := xCamEnable;

fbTabSwitch(	i_xEnable				:= (xCamEnable AND iq_stAxisModuleItf.stMultiCam.i_xEnableTabHandler),
				i_xLowEnd				:= iq_stAxisModuleItf.stMultiCam.q_xXLowEnd,
				i_xHighEnd				:= iq_stAxisModuleItf.stMultiCam.q_xXHighEnd,
				i_udiTableSelectNr		:= iq_stAxisModuleItf.stMultiCam.i_udiTableSelectNr,
				iq_xTakeNewCam			:= iq_stAxisModuleItf.stMultiCam.iq_xNewCam,
				iq_xTakeInstantNewCam	:= iq_stAxisModuleItf.stMultiCam.iq_xInstantNewCam,
				iq_xNewCam				:= xNewCam,
				iq_xInstantNewCam		:= xInstantNewCam,
				iq_astMotionPar			:= iq_stAxisModuleItf.stMultiCam.iq_astMotionPar,
				iq_stOutTab				:= stCamTab,
				q_xActive				=> ,
				q_xReady				=> ,
				q_etDiag				=> ,
				q_etDiagExt				=> ,
				q_sMsg					=> ,
				q_udiTableNumber		=> );

IF (iq_stAxisModuleItf.stMultiCam.i_udiTableSelectNr < 0) OR (iq_stAxisModuleItf.stMultiCam.i_udiTableSelectNr > AXM_GPL.Gc_udiMaxNumberOfCamTables) THEN
	iq_stAxisModuleItf.stMultiCam.i_udiTableSelectNr := 0;
ELSE
	iq_stAxisModuleItf.stMultiCam.i_udiTableSelectNr := iq_stAxisModuleItf.stMultiCam.i_udiTableSelectNr;
END_IF

IF NOT iq_stAxisModuleItf.stMultiCam.i_xEnableTabHandler THEN
	xNewCam 		:= iq_stAxisModuleItf.stMultiCam.iq_xNewCam;
	xInstantNewCam 	:= iq_stAxisModuleItf.stMultiCam.iq_xInstantNewCam;
	stCamTab 		:= iq_stAxisModuleItf.stMultiCam.iq_astMotionPar[iq_stAxisModuleItf.stMultiCam.i_udiTableSelectNr];
END_IF

fbMultiCam(	i_xEnable			:= xEnableMultiCamFb AND fbDriveEnable.q_xDriveEnabled,
			i_ifDrive			:= iq_stAxisModuleItf.stMain.i_ifDrive,
			i_xStart			:= (xStartFlag OR iq_stAxisModuleItf.stMain.i_xStart),
			i_xWsSelect			:= xWsSelect,
			i_etCsModeSlave		:= iq_stAxisModuleItf.stMultiCam.i_etCsModeSlave,
			i_etCsModeMaster	:= iq_stAxisModuleItf.stMultiCam.i_etCsModeMaster,
			i_etWsMode			:= iq_stAxisModuleItf.stMultiCam.i_etWsMode,
			i_lrWsWindow		:= iq_stAxisModuleItf.stMultiCam.i_lrWsWindow,
			i_lrWsVel			:= iq_stAxisModuleItf.stMultiCam.i_lrWsVel,
			i_lrWsAcc			:= iq_stAxisModuleItf.stMultiCam.i_lrWsAcc,
			i_lrWsJerk			:= iq_stAxisModuleItf.stMultiCam.i_lrWsJerk,
			i_xWsStart			:= xWsStartFlag,
			i_diTxEnd			:= iq_stAxisModuleItf.stMultiCam.i_diTXend,
			i_lrInstantXLimMax	:= iq_stAxisModuleItf.stMultiCam.i_lrInstantXLimMax,
 			iq_lencMaster		:= iq_stAxisModuleItf.stMain.iq_lencEncoder,
			iq_stExt			:= iq_stAxisModuleItf.stMultiCam.iq_stExt,
			iq_xNewCam			:= xNewCam,
			iq_xInstantNewCam	:= xInstantNewCam,
			iq_stMultiCamData	:= stCamTab,
			q_xActive			=> ,
			q_xReady			=> ,
			q_etDiag			=> etDiagBuffer,
			q_etDiagExt			=> etDiagExtBufferPDL,
			q_sMsg				=> sDiagMsgBuffer,
			q_xInWsWindow		=> iq_stAxisModuleItf.stMultiCam.q_xInWsWindow,
			q_xSynActive		=> iq_stAxisModuleItf.stMain.q_xSynchron,
			q_lrPositionY		=> lrCamPositionY,
			q_xXLowEnd			=> iq_stAxisModuleItf.stMultiCam.q_xXLowEnd,
			q_xXHighEnd			=> iq_stAxisModuleItf.stMultiCam.q_xXHighEnd,
			q_stActualCamData	=> iq_stAxisModuleItf.stMultiCam.q_stActualCamData);

DiagTestMultiCam(	iq_etDiag		:= fbMultiCam.q_etDiag,
					iq_etDiagExt	:= fbMultiCam.q_etDiagExt,
					iq_sMsg			:= fbMultiCam.q_sMsg);

IF (fbMultiCam.q_etDiagExt = PDL_ET_DiagExt.ShowCamPosition) THEN
	iq_stAxisModuleItf.stMultiCam.q_lrCalculatedCamPosition := lrCamPositionY;
ELSE
	iq_stAxisModuleItf.stMultiCam.q_lrCalculatedCamPosition := 0;
END_IF

IF NOT iq_stAxisModuleItf.stMultiCam.i_xEnableTabHandler THEN
	iq_stAxisModuleItf.stMultiCam.iq_xInstantNewCam := xInstantNewCam;
	iq_stAxisModuleItf.stMultiCam.iq_xNewCam 		:= xNewCam;
END_IF

IF iq_stAxisModuleItf.stMultiCam.i_xEnableTabHandler THEN
	iq_stAxisModuleItf.stMultiCam.q_diActTable := UDINT_TO_DINT(fbTabSwitch.q_udiTableNumber);
ELSE
	iq_stAxisModuleItf.stMultiCam.q_diActTable := iq_stAxisModuleItf.stMultiCam.q_stActualCamData.diUserTableId;
END_IF

IF iq_stAxisModuleItf.stMultiCam.iq_xChangeMaster THEN

	IF (iq_stAxisModuleItf.stMain.i_ifMaster = 0) THEN
		stExceptionModuleReaction2.etDiag := GD.ET_Diag.InputParameterInvalid;
		stExceptionModuleReaction2.udiDiagExt := PDL_ET_DiagExt.MasterInvalid;
		stExceptionModuleReaction2.sMsg := 'no master given';
		ReportException(iq_stException := stExceptionModuleReaction2);
	END_IF

	iq_stAxisModuleItf.stMain.iq_lencEncoder.ConnectMasterAxis(
		i_ifAxis   := iq_stAxisModuleItf.stMain.i_ifMaster,
		q_xError   => xError,
		q_etResult => etResultMoin);

	IF (iq_stAxisModuleItf.stMultiCam.i_xSetEncoderPosition) THEN
		(* set the lenc to the position of the master *)
		(* read the position of the master *)
		lrMasterPos := GetMasterPosition();

		THIS^.fbSetPos(
			Axis     := iq_stAxisModuleItf.stMain.iq_lencEncoder,
			Execute  := TRUE,
			Position := (lrMasterPos + iq_stAxisModuleItf.stMultiCam.i_lrSetEncoderOffset),
			Relative := FALSE,
			Done     =>,
			Busy     =>,
			Error    => xError,
			ErrorId  => etResultPlco);

		IF xError THEN
			stExceptionUnexpected.udiDiagExt := AXM_ET_DiagExt.UnknownFeedback;
			stExceptionUnexpected.sMsg       := Standard.CONCAT('SetEncoderPosition: ', TO_STRING(etResultPlco));
			ReportException(iq_stException := stExceptionUnexpected);
		END_IF
		THIS^.fbSetPos(Execute := FALSE);
	END_IF

	iq_stAxisModuleItf.stMultiCam.iq_xChangeMaster := FALSE;
END_IF

iq_stAxisModuleItf.stMain.q_lrPositionX := iq_stAxisModuleItf.stMain.iq_lencEncoder.lrPosition;
iq_stAxisModuleItf.stMain.q_lrPositionX := iq_stAxisModuleItf.stMain.i_ifDrive.stMotionOfMaster.lrPosition;

IF fbMultiCam.q_xReady AND NOT fbMultiCam.i_xStart
	AND NOT (fbMultiCam.q_etDiagExt = PDL_ET_DiagExt.WaitUntilStopPositionReached)
	AND NOT (fbMultiCam.q_etDiagExt = PDL_ET_DiagExt.WaitUntilCamFinished) THEN
	iq_stAxisModuleItf.stMain.q_etState := AXM_ET_State.MultiCamWaitForStart;
ELSIF fbMultiCam.q_xReady AND fbMultiCam.i_xStart AND fbMultiCam.i_xWsSelect AND NOT fbMultiCam.i_xWsStart AND NOT fbMultiCam.q_xSynActive
	AND NOT (fbMultiCam.q_etDiagExt = PDL_ET_DiagExt.ShowCamPosition) THEN
	iq_stAxisModuleItf.stMain.q_etState := AXM_ET_State.MultiCamWaitForWsStart;
ELSIF fbMultiCam.q_xReady AND fbMultiCam.i_xStart AND fbMultiCam.i_xWsSelect AND fbMultiCam.i_xWsStart AND NOT fbMultiCam.q_xSynActive THEN
	iq_stAxisModuleItf.stMain.q_etState := AXM_ET_State.MultiCamWsExecuting;
ELSIF fbMultiCam.q_xSynActive
	OR (fbMultiCam.q_etDiagExt = PDL_ET_DiagExt.ShowCamPosition)
	OR (fbMultiCam.q_etDiagExt = PDL_ET_DiagExt.WaitUntilCamStarted)
	OR (fbMultiCam.q_etDiagExt = PDL_ET_DiagExt.WaitUntilFirstCamStarted)
	OR (fbMultiCam.q_etDiagExt = PDL_ET_DiagExt.WaitForNewCam)
	OR (fbMultiCam.q_etDiagExt = PDL_ET_DiagExt.WaitUntilStopPositionReached)
	OR (fbMultiCam.q_etDiagExt = PDL_ET_DiagExt.WaitUntilCamFinished) THEN
	iq_stAxisModuleItf.stMain.q_etState := AXM_ET_State.MultiCamRunning;
ELSE
	IF xCamEnable THEN
		iq_stAxisModuleItf.stMain.q_etState := AXM_ET_State.MultiCamInit;
	ELSE
		iq_stAxisModuleItf.stMain.q_etState := AXM_ET_State.MultiCamExit;
	END_IF
END_IF

IF NOT xCamEnable AND NOT fbMultiCam.q_xActive THEN
	xCamActive := FALSE;
END_IF

(* ---- MultiCam_entry.act.st ---- *)
__METADATA__
{
  "v3Meta": {
    "objectGuid": "13a0f2e5-3dc3-4c49-bfa3-1e59ad4bbaa9",
    "objectTypeGuid": "8ac092e5-3128-4e26-9e7e-11016c6684f2",
    "embeddedObjectTypeGuids": [
      "3b83b776-fb25-43b8-99f2-3c507c9143fc"
    ],
    "properties": {},
    "subObjects": {}
  }
}

fbMultiCam.RegisterLoggerPoint(
	i_ifParent  := fbLoggerPoint,
	i_sName     := 'MultiCam',
	q_etDiag    =>,
	q_etDiagExt => );

xCamActive                          := TRUE;
iq_stAxisModuleItf.stMain.q_etState := AXM_ET_State.MultiCamInit;

IF iq_stAxisModuleItf.stMain.iq_lencEncoder = 0 THEN
	stExceptionModuleReaction2.etDiag     := GD.ET_Diag.InputParameterInvalid;
	stExceptionModuleReaction2.udiDiagExt := AXM_ET_DiagExt.LencInvalid;
	stExceptionModuleReaction2.sMsg       := 'No logical Encoder connected on input iq_lencEncoder';
	ReportException(iq_stException := stExceptionModuleReaction2);
ELSIF iq_stAxisModuleItf.stMain.iq_lencEncoder.xIsModulo AND iq_stAxisModuleItf.stMultiCam.i_xCheckEncoderPeriod THEN
	stExceptionModuleReaction2.etDiag     := GD.ET_Diag.InputParameterInvalid;
	stExceptionModuleReaction2.udiDiagExt := AXM_ET_DiagExt.PeriodRange;
	stExceptionModuleReaction2.sMsg       := 'Lenc is set to Modulo';
	ReportException(iq_stException := stExceptionModuleReaction2);
ELSIF (iq_stAxisModuleItf.stMain.i_ifMaster = 0) THEN
	stExceptionModuleReaction2.etDiag     := GD.ET_Diag.InputParameterInvalid;
	stExceptionModuleReaction2.udiDiagExt := AXM_ET_DiagExt.MasterInvalid;
	stExceptionModuleReaction2.sMsg       := 'no master given';
	ReportException(iq_stException := stExceptionModuleReaction2);
ELSE
	//replace of FC_SetMasterEncoder
	iq_stAxisModuleItf.stMain.iq_lencEncoder.ConnectMasterAxis(
		i_ifAxis   := iq_stAxisModuleItf.stMain.i_ifMaster,
		q_xError   => xError,
		q_etResult => etResultMoin);

	IF xError THEN
		stExceptionUnexpected.udiDiagExt := AXM_ET_DiagExt.MasterInvalid;
		stExceptionUnexpected.sMsg       := TO_STRING(etResultMoin);
		ReportException(iq_stException := stExceptionUnexpected);
	END_IF

	IF (iq_stAxisModuleItf.stMultiCam.i_xSetEncoderPosition) THEN
		(* set the lenc to the position of the master *)
		(* read the position of the master *)
		lrMasterPos := GetMasterPosition();

		THIS^.fbSetPos(
			Axis     := iq_stAxisModuleItf.stMain.iq_lencEncoder,
			Execute  := TRUE,
			Position := (lrMasterPos + iq_stAxisModuleItf.stMultiCam.i_lrSetEncoderOffset),
			Relative := FALSE,
			Done     =>,
			Busy     =>,
			Error    => xError,
			ErrorId  => etResultPlco);

		IF xError THEN
			stExceptionUnexpected.udiDiagExt := AXM_ET_DiagExt.UnknownFeedback;
			stExceptionUnexpected.sMsg       := Standard.CONCAT('SetEncoderPosition: ', TO_STRING(etResultPlco));
			ReportException(iq_stException := stExceptionUnexpected);
		END_IF
	END_IF
END_IF

THIS^.fbSetPos(Execute := FALSE);
iq_stAxisModuleItf.stMain.q_lrPositionX := iq_stAxisModuleItf.stMain.i_ifDrive.stMotionOfMaster.lrPosition;

(* ---- MultiCam_exit.act.st ---- *)
__METADATA__
{
  "v3Meta": {
    "objectGuid": "05cae1eb-9684-4632-bef6-8a05e37eeba1",
    "objectTypeGuid": "8ac092e5-3128-4e26-9e7e-11016c6684f2",
    "embeddedObjectTypeGuids": [
      "3b83b776-fb25-43b8-99f2-3c507c9143fc"
    ],
    "properties": {},
    "subObjects": {}
  }
}

(* Disconnection *)
IF NOT iq_stAxisModuleItf.stMultiCam.i_xKeepEncoderConnection THEN
	iq_stAxisModuleItf.stMain.iq_lencEncoder.DisconnectMasterAxis(
									q_xError 	=> xError,
									q_etResult  => etResultMoin);

	IF xError THEN
		stExceptionUnexpected.udiDiagExt := AXM_ET_DiagExt.UnknownFeedback;
		stExceptionUnexpected.sMsg := TO_STRING(etResultMoin);
		ReportException(iq_stException := stExceptionUnexpected);
	END_IF

END_IF
iq_stAxisModuleItf.stMain.q_lrPositionX := 0.0;

(* ---- NoOp_active.act.st ---- *)
__METADATA__
{
  "v3Meta": {
    "objectGuid": "30bfc610-6151-43e5-88b1-85d38d3fc0ea",
    "objectTypeGuid": "8ac092e5-3128-4e26-9e7e-11016c6684f2",
    "embeddedObjectTypeGuids": [
      "3b83b776-fb25-43b8-99f2-3c507c9143fc"
    ],
    "properties": {},
    "subObjects": {}
  }
}

iq_stAxisModuleItf.stMain.q_etOpMode := AXM_ET_OpMode.NoOp;
IF fbDriveEnable.q_xDriveEnabled THEN
	iq_stAxisModuleItf.stMain.q_etState := AXM_ET_State.NoOpDriveEnabled;
ELSE
	iq_stAxisModuleItf.stMain.q_etState := AXM_ET_State.NoOpDriveDisabled;
END_IF

(* ---- Output_active.act.st ---- *)
__METADATA__
{
  "v3Meta": {
    "objectGuid": "e6be1b92-6fa1-4507-8656-3f00fb93657e",
    "objectTypeGuid": "8ac092e5-3128-4e26-9e7e-11016c6684f2",
    "embeddedObjectTypeGuids": [
      "3b83b776-fb25-43b8-99f2-3c507c9143fc"
    ],
    "properties": {},
    "subObjects": {}
  }
}

IF xNotAbleToSetException THEN
	; (* Do nothing. Diag outputs show not reportable exception *)
	iq_stStandardModuleItf.q_xReady := FALSE;
ELSIF stModuleReaction.axReaction[TPL.ET_Reaction.AsyncStop] THEN
	iq_stStandardModuleItf.q_etDiag := GD.ET_Diag.ExecutionAborted;
	iq_stStandardModuleItf.q_udiDiagExt := AXM_ET_DiagExt.AsyncStop;
	iq_stStandardModuleItf.q_sDiagExt := 'AsyncStop';
	iq_stStandardModuleItf.q_sMsg := AXM_FC_EtDiagExtToString(i_etDiagExt := AXM_ET_DiagExt.AsyncStop);
	iq_stStandardModuleItf.q_xReady := FALSE;
ELSIF stModuleReaction.axReaction[TPL.ET_Reaction.SyncStopEL] THEN
	iq_stStandardModuleItf.q_etDiag := GD.ET_Diag.ExecutionAborted;
	iq_stStandardModuleItf.q_udiDiagExt := AXM_ET_DiagExt.SyncStopEL;
	iq_stStandardModuleItf.q_sDiagExt := 'SyncStopEL';
	iq_stStandardModuleItf.q_sMsg := AXM_FC_EtDiagExtToString(i_etDiagExt := AXM_ET_DiagExt.SyncStopEL);
	iq_stStandardModuleItf.q_xReady := FALSE;
ELSIF stModuleReaction.axReaction[TPL.ET_Reaction.SyncStopEH] THEN
	iq_stStandardModuleItf.q_etDiag := GD.ET_Diag.ExecutionAborted;
	iq_stStandardModuleItf.q_udiDiagExt := AXM_ET_DiagExt.SyncStopEH;
	iq_stStandardModuleItf.q_sDiagExt := 'SyncStopEH';
	iq_stStandardModuleItf.q_sMsg := AXM_FC_EtDiagExtToString(i_etDiagExt := AXM_ET_DiagExt.SyncStopEH);
	iq_stStandardModuleItf.q_xReady := FALSE;
ELSIF stModuleReaction.axReaction[TPL.ET_Reaction.StopEndOfCycle] THEN
	iq_stStandardModuleItf.q_etDiag := GD.ET_Diag.ExecutionAborted;
	iq_stStandardModuleItf.q_udiDiagExt := AXM_ET_DiagExt.StopEndOfCycle;
	iq_stStandardModuleItf.q_sDiagExt := 'StopEndOfCycle';
	iq_stStandardModuleItf.q_sMsg := AXM_FC_EtDiagExtToString(i_etDiagExt := AXM_ET_DiagExt.StopEndOfCycle);
	iq_stStandardModuleItf.q_xReady := FALSE;
ELSE
	IF (iq_stStandardModuleItf.i_xEnable) AND
		(iq_stAxisModuleItf.stMain.q_etState <> AXM_ET_State.Disabled) AND
		(iq_stAxisModuleItf.stMain.q_etState <> AXM_ET_State.Initializing) THEN
		iq_stStandardModuleItf.q_xReady := TRUE;
	ELSE
		iq_stStandardModuleItf.q_xReady := FALSE;
	END_IF
	iq_stStandardModuleItf.q_etDiag := GD.ET_Diag.Ok;
	CASE iq_stAxisModuleItf.stMain.q_etState OF
		AXM_ET_State.Disabled:
			iq_stStandardModuleItf.q_udiDiagExt := AXM_ET_DiagExt.Disabled;
		AXM_ET_State.Initializing:
			iq_stStandardModuleItf.q_udiDiagExt := AXM_ET_DiagExt.Initializing;
		AXM_ET_State.NoOpDriveEnabled:
			iq_stStandardModuleItf.q_udiDiagExt := AXM_ET_DiagExt.NoOpDriveEnabled;
		AXM_ET_State.NoOpDriveDisabled:
			iq_stStandardModuleItf.q_udiDiagExt := AXM_ET_DiagExt.NoOpDriveDisabled;
		AXM_ET_State.HomingInit:
			iq_stStandardModuleItf.q_udiDiagExt := AXM_ET_DiagExt.HomingInit;
		AXM_ET_State.HomingWaitForStart:
			iq_stStandardModuleItf.q_udiDiagExt := AXM_ET_DiagExt.HomingWaitForStart;
		AXM_ET_State.HomingExecuting:
			iq_stStandardModuleItf.q_udiDiagExt := AXM_ET_DiagExt.HomingExecuting;
		AXM_ET_State.HomingDone:
			iq_stStandardModuleItf.q_udiDiagExt := AXM_ET_DiagExt.HomingDone;
		AXM_ET_State.HomingExit:
			iq_stStandardModuleItf.q_udiDiagExt := AXM_ET_DiagExt.HomingExit;
		AXM_ET_State.ManualInit:
			iq_stStandardModuleItf.q_udiDiagExt := AXM_ET_DiagExt.ManualInit;
		AXM_ET_State.ManualRunning:
			iq_stStandardModuleItf.q_udiDiagExt := AXM_ET_DiagExt.ManualRunning;
		AXM_ET_State.ManualExit:
			iq_stStandardModuleItf.q_udiDiagExt := AXM_ET_DiagExt.ManualExit;
		AXM_ET_State.MultiCamInit:
			iq_stStandardModuleItf.q_udiDiagExt := AXM_ET_DiagExt.MultiCamInit;
		AXM_ET_State.MultiCamWaitForStart:
			iq_stStandardModuleItf.q_udiDiagExt := AXM_ET_DiagExt.MultiCamWaitForStart;
		AXM_ET_State.MultiCamWaitForWsStart:
			iq_stStandardModuleItf.q_udiDiagExt := AXM_ET_DiagExt.MultiCamWaitForWsStart;
		AXM_ET_State.MultiCamWsExecuting:
			iq_stStandardModuleItf.q_udiDiagExt := AXM_ET_DiagExt.MultiCamWsExecuting;
		AXM_ET_State.MultiCamRunning:
			iq_stStandardModuleItf.q_udiDiagExt := AXM_ET_DiagExt.MultiCamRunning;
		AXM_ET_State.MultiCamExit:
			iq_stStandardModuleItf.q_udiDiagExt := AXM_ET_DiagExt.MultiCamExit;
		AXM_ET_State.EndlessInit:
			iq_stStandardModuleItf.q_udiDiagExt := AXM_ET_DiagExt.EndlessInit;
		AXM_ET_State.EndlessWaitForStart:
			iq_stStandardModuleItf.q_udiDiagExt := AXM_ET_DiagExt.EndlessWaitForStart;
		AXM_ET_State.EndlessRunning:
			iq_stStandardModuleItf.q_udiDiagExt := AXM_ET_DiagExt.EndlessRunning;
		AXM_ET_State.EndlessExit:
			iq_stStandardModuleItf.q_udiDiagExt := AXM_ET_DiagExt.EndlessExit;
		AXM_ET_State.PositioningInit:
			iq_stStandardModuleItf.q_udiDiagExt := AXM_ET_DiagExt.PositioningInit;
		AXM_ET_State.PositioningWaitForStart:
			iq_stStandardModuleItf.q_udiDiagExt := AXM_ET_DiagExt.PositioningWaitForStart;
		AXM_ET_State.PositioningRunning:
			iq_stStandardModuleItf.q_udiDiagExt := AXM_ET_DiagExt.PositioningRunning;
		AXM_ET_State.PositioningExit:
			iq_stStandardModuleItf.q_udiDiagExt := AXM_ET_DiagExt.PositioningExit;
		AXM_ET_State.BrakeReleaseInit:
			iq_stStandardModuleItf.q_udiDiagExt := AXM_ET_DiagExt.BrakeReleaseInit;
		AXM_ET_State.BrakeClosed:
			iq_stStandardModuleItf.q_udiDiagExt := AXM_ET_DiagExt.BrakeClosed;
		AXM_ET_State.BrakeReleased:
			iq_stStandardModuleItf.q_udiDiagExt := AXM_ET_DiagExt.BrakeReleased;
		AXM_ET_State.BrakeReleaseExit:
			iq_stStandardModuleItf.q_udiDiagExt := AXM_ET_DiagExt.BrakeReleaseExit;
		AXM_ET_State.AdditionalInit:
			iq_stStandardModuleItf.q_udiDiagExt := AXM_ET_DiagExt.AdditionalInit;
		AXM_ET_State.AdditionalWaitForStart:
			iq_stStandardModuleItf.q_udiDiagExt := AXM_ET_DiagExt.AdditionalWaitForStart;
		AXM_ET_State.AdditionalRunning:
			iq_stStandardModuleItf.q_udiDiagExt := AXM_ET_DiagExt.AdditionalRunning;
		AXM_ET_State.AdditionalExit:
			iq_stStandardModuleItf.q_udiDiagExt := AXM_ET_DiagExt.AdditionalExit;
	END_CASE
	iq_stStandardModuleItf.q_sDiagExt := AXM_FC_EtDiagExtToString(i_etDiagExt := iq_stStandardModuleItf.q_udiDiagExt);
	iq_stStandardModuleItf.q_sMsg := AXM_FC_EtDiagExtToString(i_etDiagExt := iq_stStandardModuleItf.q_udiDiagExt);
END_IF

IF iq_stStandardModuleItf.q_xActive THEN
	iq_stAxisModuleItf.stMain.q_lrPosition := iq_stAxisModuleItf.stMain.i_ifDrive.lrPosition;
ELSE
	iq_stStandardModuleItf.q_xException := FALSE;
	xInitActualValuesPos := FALSE;
END_IF

IF fbLoggerPoint.etLogLevel >= APL.ET_LogLevel.StatusMessage THEN
	IF (iq_stAxisModuleItf.stMain.q_etOpMode <> etOpModeOld) THEN
		fbLoggerPoint.AddLogEntry(	i_etLogLevel	:= APL.ET_LogLevel.StatusMessage,
									i_etDiag		:= GD.ET_Diag.Ok,
									i_udiDiagExt	:= AXM_ET_DiagExt.Ok,
									i_sMessage		:= Standard.CONCAT('OpMode changed to: ', AXM_FC_EtOpModeToString(i_etOpMode := iq_stAxisModuleItf.stMain.q_etOpMode)),
									q_etDiag		:= ,
									q_etDiagExt		:= );
	END_IF
	etOpModeOld := iq_stAxisModuleItf.stMain.q_etOpMode;

	IF (iq_stAxisModuleItf.stMain.q_etState <> etStateOld) THEN
		fbLoggerPoint.AddLogEntry(	i_etLogLevel	:= APL.ET_LogLevel.StatusMessage,
									i_etDiag		:= GD.ET_Diag.Ok,
									i_udiDiagExt	:= AXM_ET_DiagExt.Ok,
									i_sMessage		:= Standard.CONCAT('State changed to: ', AXM_FC_EtStateToString(i_etState := iq_stAxisModuleItf.stMain.q_etState)),
									q_etDiag		:= ,
									q_etDiagExt		:= );
	END_IF
	etStateOld := iq_stAxisModuleItf.stMain.q_etState;
END_IF

(* ---- Positioning_active.act.st ---- *)
__METADATA__
{
  "v3Meta": {
    "objectGuid": "2ecf66ce-f923-48fb-8d77-3fe74e91c2a1",
    "objectTypeGuid": "8ac092e5-3128-4e26-9e7e-11016c6684f2",
    "embeddedObjectTypeGuids": [
      "3b83b776-fb25-43b8-99f2-3c507c9143fc"
    ],
    "properties": {},
    "subObjects": {}
  }
}

iq_stAxisModuleItf.stMain.q_etOpMode := AXM_ET_OpMode.Positioning;

IF (iq_stAxisModuleItf.stMain.stReducedVelocity.i_xEnableReducedVelocity AND
	NOT iq_stAxisModuleItf.stMain.stReducedVelocity.i_xOnlyLimitCheck) THEN

	lrPosVel := MIN(iq_stAxisModuleItf.stPos.i_lrVel, iq_stAxisModuleItf.stMain.stReducedVelocity.i_lrMaxReducedVelocity);
ELSE
	lrPosVel := iq_stAxisModuleItf.stPos.i_lrVel;
END_IF

lrPosVel := iq_stAxisModuleItf.stPos.i_lrVel;

IF iq_stAxisModuleItf.stPos.i_xStop THEN
	xStartFlag := FALSE;
END_IF
xPosStart := (xStartFlag OR iq_stAxisModuleItf.stMain.i_xStart) AND NOT stModuleReaction.axReaction[TPL.ET_Reaction.StopEndOfCycle];

fbVarioPos(
	i_xEnable                  := xPosEnable AND fbDriveEnable.q_xDriveEnabled,
	i_ifDrive                  := iq_stAxisModuleItf.stMain.i_ifDrive,
	i_xStart                   := xPosStart,
	i_xStop                    := iq_stAxisModuleItf.stPos.i_xStop,
	i_lrTarget                 := iq_stAxisModuleItf.stPos.i_lrTarget,
	i_lrVel                    := lrPosVel,
	i_lrAcc                    := iq_stAxisModuleItf.stPos.i_lrAcc,
	i_lrDec                    := iq_stAxisModuleItf.stPos.i_lrDec,
	i_lrJerk                   := iq_stAxisModuleItf.stPos.i_lrJerk,
	i_etPosMode                := iq_stAxisModuleItf.stPos.i_etPosMode,
	q_xActive                  => xPosActive,
	q_xReady                   =>,
	q_etDiag                   => etDiagBuffer,
	q_etDiagExt                => etDiagExtBufferPDL,
	q_sMsg                     => sDiagMsgBuffer,
	q_xMotionInstructionActive =>,
	q_lrPosition               =>,
	q_xInPosition              => iq_stAxisModuleItf.stPos.q_xInPosition);

DiagTestPositioning(
	iq_etDiag    := fbVarioPos.q_etDiag,
	iq_etDiagExt := fbVarioPos.q_etDiagExt,
	iq_sMsg      := fbVarioPos.q_sMsg);

IF fbVarioPos.q_xReady AND NOT fbVarioPos.q_xMotionInstructionActive THEN
	iq_stAxisModuleItf.stMain.q_etState := AXM_ET_State.PositioningWaitForStart;
ELSIF fbVarioPos.q_xReady AND fbVarioPos.q_xMotionInstructionActive THEN
	iq_stAxisModuleItf.stMain.q_etState := AXM_ET_State.PositioningRunning;
ELSE
	IF xPosEnable THEN
		iq_stAxisModuleItf.stMain.q_etState := AXM_ET_State.PositioningInit;
	ELSE
		iq_stAxisModuleItf.stMain.q_etState := AXM_ET_State.PositioningExit;
	END_IF
END_IF

(* make shure next start command is effective *)
IF fbVarioPos.q_xMotionInstructionActive AND xMotionActiveOld THEN
	xStartFlag := FALSE;
END_IF
xMotionActiveOld := fbVarioPos.q_xMotionInstructionActive;

IF NOT xPosEnable AND NOT fbVarioPos.q_xActive THEN
	xPosActive := FALSE;
END_IF

(* ---- PowerControl_active.act.st ---- *)
__METADATA__
{
  "v3Meta": {
    "objectGuid": "3ace14da-dde1-48a4-ba04-45999c630589",
    "objectTypeGuid": "8ac092e5-3128-4e26-9e7e-11016c6684f2",
    "embeddedObjectTypeGuids": [
      "3b83b776-fb25-43b8-99f2-3c507c9143fc"
    ],
    "properties": {},
    "subObjects": {}
  }
}

(* ------------------------------------------------------------------------------------------------------------------------------------------------------*)
(* Controller State Machine *)
(* ------------------------------------------------------------------------------------------------------------------------------------------------------*)

CASE etPowerState OF

	AXM_ET_PowerState.Disabled:	(* Error or Disabled *)
		;

(* ------------------------------------------------------------------------------------------------------------------------------------------------------*)
	AXM_ET_PowerState.PowerOff:	(* Controller State: Axis disabled, wait for PowerOn *)
(* ------------------------------------------------------------------------------------------------------------------------------------------------------*)
		fbDriveEnable(	i_xEnable		:= TRUE,
						i_ifDrive		:= iq_stAxisModuleItf.stMain.i_ifDrive,
						i_xEnableDrive	:= xCMDPowerOn AND NOT fbHome.q_xDisableDrive,
						i_xDiagQuit		:= iq_stStandardModuleItf.i_xDiagQuit,
						q_xActive		=> ,
						q_xReady		=> ,
						q_etDiag		=> etDiagBuffer,
						q_etDiagExt		=> etDiagExtBufferPDL,
						q_sMsg			=> sDiagMsgBuffer,
						q_xDriveEnabled	=> );
		IF (etDiagBuffer <> GD.ET_Diag.Ok) THEN
			DiagTestDriveEnable(	iq_etDiag		:= fbDriveEnable.q_etDiag,
									iq_etDiagExt	:= fbDriveEnable.q_etDiagExt,
									iq_sMsg			:= fbDriveEnable.q_sMsg);
		ELSIF fbDriveEnable.q_xDriveEnabled THEN
			etPowerState := AXM_ET_PowerState.PowerOn;
		END_IF

(* ------------------------------------------------------------------------------------------------------------------------------------------------------*)
	AXM_ET_PowerState.PowerOn:	(* Controller State: AxisEnabled, wait for PowerOff  *)
(* ------------------------------------------------------------------------------------------------------------------------------------------------------*)
		fbDriveEnable(	i_xEnable		:= TRUE,
						i_ifDrive		:= iq_stAxisModuleItf.stMain.i_ifDrive,
						i_xEnableDrive	:= xCMDPowerOn AND NOT fbHome.q_xDisableDrive,
						i_xDiagQuit		:= iq_stStandardModuleItf.i_xDiagQuit,
						q_xActive		=> ,
						q_xReady		=> ,
						q_etDiag		=> etDiagBuffer,
						q_etDiagExt		=> etDiagExtBufferPDL,
						q_sMsg			=> sDiagMsgBuffer,
						q_xDriveEnabled	=> );
		IF (etDiagBuffer <> GD.ET_Diag.Ok) THEN
			DiagTestDriveEnable(	iq_etDiag		:= fbDriveEnable.q_etDiag,
									iq_etDiagExt	:= fbDriveEnable.q_etDiagExt,
									iq_sMsg			:= fbDriveEnable.q_sMsg);
		ELSIF NOT fbDriveEnable.q_xDriveEnabled THEN
			etPowerState := AXM_ET_PowerState.PowerOff;
		END_IF

(* ------------------------------------------------------------------------------------------------------------------------------------------------------*)
	AXM_ET_PowerState.WaitForDisabled:   (* Controller State: wait for FB_Axis_Enable  not active  *)
(* ------------------------------------------------------------------------------------------------------------------------------------------------------*)
		fbDriveEnable(	i_xEnable		:= FALSE,
						i_ifDrive		:= iq_stAxisModuleItf.stMain.i_ifDrive,
						i_xEnableDrive	:= FALSE,
						i_xDiagQuit		:= FALSE,
						q_xActive		=> ,
						q_xReady		=> ,
						q_etDiag		=> etDiagBuffer,
						q_etDiagExt		=> etDiagExtBufferPDL,
						q_sMsg			=> sDiagMsgBuffer,
						q_xDriveEnabled	=> );

		IF (etDiagBuffer <> GD.ET_Diag.Ok) THEN
			DiagTestDriveEnable(	iq_etDiag		:= fbDriveEnable.q_etDiag,
									iq_etDiagExt	:= fbDriveEnable.q_etDiagExt,
									iq_sMsg			:= fbDriveEnable.q_sMsg);
		ELSIF NOT fbDriveEnable.q_xActive THEN
			etPowerState := AXM_ET_PowerState.Disabled;
			iq_stAxisModuleItf.stMain.q_etState := AXM_ET_State.NoOpDriveDisabled;
		END_IF
END_CASE

IF	(iq_stAxisModuleItf.stMain.i_ifDrive.etAxisState > MOIN.ET_AxisState.Disabled) THEN
	iq_stAxisModuleItf.stMain.q_xDriveActive := TRUE;
ELSE
	iq_stAxisModuleItf.stMain.q_xDriveActive := FALSE;
END_IF

(********************** xMotionActive ************************)
IF (iq_stAxisModuleItf.stMain.i_lrMotionActiveVelLimit < 0) THEN
	stExceptionModuleReaction3.etDiag := GD.ET_Diag.InputParameterInvalid;
	stExceptionModuleReaction3.udiDiagExt := AXM_ET_DiagExt.MotionActiveVelLimitRange;
	stExceptionModuleReaction3.sMsg := 'has to be >= 0';
	ReportException(iq_stException := stExceptionModuleReaction3);
ELSE
	GetInterfaces();
	IF iq_stAxisModuleItf.stMain.i_etMotionActiveVelType = AXM_ET_MotionActiveVelType.RefVelocity
		OR iq_stAxisModuleItf.stMain.i_etMotionActiveVelType = AXM_ET_MotionActiveVelType.MechRefVelocity
	THEN
		iq_stAxisModuleItf.stMain.q_xMotionActive := ( ABS(iq_stAxisModuleItf.stMain.i_ifDrive.RefVelocity) > iq_stAxisModuleItf.stMain.i_lrMotionActiveVelLimit);

	ELSIF iq_stAxisModuleItf.stMain.i_etMotionActiveVelType = AXM_ET_MotionActiveVelType.MechVelocity
		OR iq_stAxisModuleItf.stMain.i_etMotionActiveVelType = AXM_ET_MotionActiveVelType.Velocity
	THEN
		iq_stAxisModuleItf.stMain.q_xMotionActive := ( ABS(ifDrive.ActualVelocity) > iq_stAxisModuleItf.stMain.i_lrMotionActiveVelLimit);
	END_IF

END_IF

(* ---- ReadTrackingDeviation.meth.st ---- *)
METHOD ReadTrackingDeviation : LREAL

VAR_OUTPUT
	q_sLrealConversion	: STRING[80];
END_VAR
VAR
	etConversionDiag	: SE_CTBX.ET_Result;
END_VAR

	GetInterfaces();

	IF ifDrive2 <> 0 THEN
		ReadTrackingDeviation :=  ifDrive2.TrackingDeviation;

		q_sLrealConversion := SE_CTBX.FC_LrealToString(
									i_sFormat := '10#0.______',
									i_lrInput := ReadTrackingDeviation,
									q_etResult => etConversionDiag,
									q_sResultMsg =>
									);

		IF etConversionDiag <> SE_CTBX.ET_Result.Ok THEN
			q_sLrealConversion := 'LREAL too big';
		END_IF
	ELSE
		q_sLrealConversion := 'TrackingDeviation not available';
		ReadTrackingDeviation := 0.0;
	END_IF

(* ---- RefuseCommand.meth.st ---- *)
{attribute 'conditionalshow_all_locals'}
METHOD INTERNAL RefuseCommand
VAR_INPUT
END_VAR

iq_stStandardModuleItf.q_xCmdActive := FALSE;
iq_stStandardModuleItf.q_xCmdDone := FALSE;
iq_stStandardModuleItf.iq_diCMD := -iq_stStandardModuleItf.iq_diCMD;

xCommandRefused := TRUE;

(* ---- RegisterLoggerPoint.meth.st ---- *)
{attribute 'conditionalshow_all_locals'}
METHOD PUBLIC RegisterLoggerPoint
VAR_INPUT
	i_ifParent		: APL.IF_LoggerPoint;
	i_sName			: STRING[80];
END_VAR
VAR_OUTPUT
	q_etDiag		: GD.ET_Diag := GD.ET_Diag.Ok;
	q_etDiagExt		: AXM_ET_DiagExt := AXM_ET_DiagExt.Ok;
END_VAR
VAR
	etDiagBuffer		: GD.ET_Diag;
	etDiagExtBufferAPL	: APL.ET_DiagExt;
END_VAR

THIS^.fbLoggerPoint.RegisterLoggerPoint(	i_ifParent		:= i_ifParent,
											i_sName			:= i_sName,
											i_sType			:= 'FB_AxisModule',
											i_sSource		:= 'AXM',
											q_etDiag		=> etDiagBuffer,
											q_etDiagExt		=> etDiagExtBufferAPL);
IF (etDiagBuffer <> GD.ET_Diag.Ok) THEN
	CASE etDiagExtBufferAPL OF
		APL.ET_DiagExt.ParentInvalid:
			q_etDiag := GD.ET_Diag.InputParameterInvalid;
			q_etDiagExt := AXM_ET_DiagExt.ParentInvalid;

		APL.ET_DiagExt.ParentNotRegistered:
			q_etDiag := GD.ET_Diag.InputParameterInvalid;
			q_etDiagExt := AXM_ET_DiagExt.ParentNotRegistered;

		APL.ET_DiagExt.MaxNumberOfLoggerPointsExeeded:
			q_etDiag := GD.ET_Diag.InputParameterInvalid;
			q_etDiagExt := AXM_ET_DiagExt.MaxNumberOfLoggerPointsExeeded;

	ELSE
		q_etDiag := GD.ET_Diag.UnexpectedProgramBehavior;
		q_etdiagExt := AXM_ET_DiagExt.UnexpectedDiagExt;
	END_CASE
END_IF

(* ---- ReportException.meth.st ---- *)
METHOD ReportException
VAR_IN_OUT
	iq_stException	: TPL.ST_Exception;
END_VAR
VAR CONSTANT
	c_diMaxReaction	: DINT := 4;
END_VAR

IF (fbLoggerPoint.etLogLevel >= APL.ET_LogLevel.CriticalException) AND (iq_stException.etDiag = GD.ET_Diag.UnexpectedProgramBehavior) THEN
	IF NOT TPL.FC_CheckExceptionIsInList( iq_stException := iq_stException, iq_stExceptionList := THIS^.iq_stExceptionList) THEN
		fbLoggerPoint.AddLogEntry(	i_etLogLevel	:= APL.ET_LogLevel.CriticalException,
									i_etDiag		:= GD.ET_Diag.Ok,
									i_udiDiagExt	:= AXM_ET_DiagExt.Ok,
									i_sMessage		:= Standard.CONCAT(Standard.CONCAT(Standard.CONCAT(Standard.CONCAT(Standard.CONCAT(Standard.CONCAT('Exception ET_Diag: ',GD.FC_EtDiagToString(i_etDiag := iq_stException.etDiag)),' ET_DiagExt: '),AXM_FC_EtDiagExtToString(i_etDiagExt := iq_stException.udiDiagExt)),' sMsg: '),iq_stException.sMsg),TPL.FC_GetStandardReactionName(iq_stReaction := iq_stException.stReaction)),
									q_etDiag		:= ,
									q_etDiagExt		:= );
	END_IF
ELSIF (fbLoggerPoint.etLogLevel >= APL.ET_LogLevel.Exception) THEN
	IF NOT TPL.FC_CheckExceptionIsInList( iq_stException := iq_stException, iq_stExceptionList := THIS^.iq_stExceptionList) THEN
		fbLoggerPoint.AddLogEntry(	i_etLogLevel	:= APL.ET_LogLevel.Exception,
									i_etDiag		:= GD.ET_Diag.Ok,
									i_udiDiagExt	:= AXM_ET_DiagExt.Ok,
									i_sMessage		:= Standard.CONCAT(Standard.CONCAT(Standard.CONCAT(Standard.CONCAT(Standard.CONCAT(Standard.CONCAT('Exception ET_Diag: ',GD.FC_EtDiagToString(i_etDiag := iq_stException.etDiag)),' ET_DiagExt: '),AXM_FC_EtDiagExtToString(i_etDiagExt := iq_stException.udiDiagExt)),' sMsg: '),iq_stException.sMsg),TPL.FC_GetStandardReactionName(iq_stReaction := iq_stException.stReaction)),
									q_etDiag		:= ,
									q_etDiagExt		:= );
	END_IF
END_IF

iq_stException.sDiagExt := AXM_FC_EtDiagExtToString(i_etDiagExt := iq_stException.udiDiagExt);
TPL.FC_SetException(	i_xExceptionActive	:= TRUE,
						iq_stException		:= iq_stException,
						iq_stExceptionList	:= iq_stExceptionList,
						iq_stLogDataList	:= iq_stLogDataList,
						q_etDiag 			=> etDiagBuffer,
						q_etDiagExt 		=> etDiagExtBufferTPL,
						q_sMsg 				=> sDiagMsgBuffer);
IF (etDiagBuffer <> GD.ET_Diag.Ok) THEN
	(* if exception could not be reported, show exception on outputs *)
	xNotAbleToSetException := TRUE;
	iq_stStandardModuleItf.q_etDiag := iq_stException.etDiag;
	iq_stStandardModuleItf.q_udiDiagExt := iq_stException.udiDiagExt;
	iq_stStandardModuleItf.q_sDiagExt := iq_stException.sDiagExt;
	iq_stStandardModuleItf.q_sMsg := iq_stException.sMsg;
END_IF

iq_stStandardModuleItf.q_xException := TRUE;

stLocalReaction.axReaction[TPL.ET_Reaction.MainsContactorOff] := stLocalReaction.axReaction[TPL.ET_Reaction.MainsContactorOff] OR iq_stException.stReaction.axReaction[iq_stStandardModuleItf.iq_stExt.udiReactionOffset + TPL.ET_Reaction.MainsContactorOff];
stLocalReaction.axReaction[TPL.ET_Reaction.AsyncStop] := stLocalReaction.axReaction[TPL.ET_Reaction.AsyncStop] OR iq_stException.stReaction.axReaction[iq_stStandardModuleItf.iq_stExt.udiReactionOffset + TPL.ET_Reaction.AsyncStop];
stLocalReaction.axReaction[TPL.ET_Reaction.SyncStopEH] := stLocalReaction.axReaction[TPL.ET_Reaction.SyncStopEH] OR iq_stException.stReaction.axReaction[iq_stStandardModuleItf.iq_stExt.udiReactionOffset + TPL.ET_Reaction.SyncStopEH];
stLocalReaction.axReaction[TPL.ET_Reaction.SyncStopEL] := stLocalReaction.axReaction[TPL.ET_Reaction.SyncStopEL] OR iq_stException.stReaction.axReaction[iq_stStandardModuleItf.iq_stExt.udiReactionOffset + TPL.ET_Reaction.SyncStopEL];
(* special handling for StopEndOfCycle. Wait till reaction feedback from machine. User can transform this reaction and make own reaction.
stLocalReaction.axReaction[TPL.ET_Reaction.StopEndOfCycle] := stLocalReaction.axReaction[TPL.ET_Reaction.StopEndOfCycle] OR iq_stException.stReaction.axReaction[TPL.ET_Reaction.StopEndOfCycle];
*)

stModuleReaction.axReaction[TPL.ET_Reaction.MainsContactorOff] := stModuleReaction.axReaction[TPL.ET_Reaction.MainsContactorOff] OR iq_stException.stReaction.axReaction[iq_stStandardModuleItf.iq_stExt.udiReactionOffset + TPL.ET_Reaction.MainsContactorOff];
stModuleReaction.axReaction[TPL.ET_Reaction.AsyncStop] := stModuleReaction.axReaction[TPL.ET_Reaction.AsyncStop] OR iq_stException.stReaction.axReaction[iq_stStandardModuleItf.iq_stExt.udiReactionOffset + TPL.ET_Reaction.AsyncStop];
stModuleReaction.axReaction[TPL.ET_Reaction.SyncStopEH] := stModuleReaction.axReaction[TPL.ET_Reaction.SyncStopEH]OR iq_stException.stReaction.axReaction[iq_stStandardModuleItf.iq_stExt.udiReactionOffset + TPL.ET_Reaction.SyncStopEH];
stModuleReaction.axReaction[TPL.ET_Reaction.SyncStopEL] := stModuleReaction.axReaction[TPL.ET_Reaction.SyncStopEL] OR iq_stException.stReaction.axReaction[iq_stStandardModuleItf.iq_stExt.udiReactionOffset + TPL.ET_Reaction.SyncStopEL];
(* special handling for StopEndOfCycle. Wait till reaction feedback from machine. User can transform this reaction and make own reaction.
stModuleReaction.axReaction[TPL.ET_Reaction.StopEndOfCycle] := stModuleReaction.axReaction[TPL.ET_Reaction.StopEndOfCycle] OR iq_stException.stReaction.axReaction[iq_stStandardModuleItf.iq_stExt.udiReactionOffset + TPL.ET_Reaction.StopEndOfCycle];
*)

(* ---- SignalSuccessfulExecution.meth.st ---- *)
{attribute 'conditionalshow_all_locals'}
METHOD INTERNAL SignalSuccessfulExecution
VAR_INPUT
END_VAR

IF fbLoggerPoint.etLogLevel >= APL.ET_LogLevel.StatusMessage THEN
	fbLoggerPoint.AddLogEntry(	i_etLogLevel	:= APL.ET_LogLevel.StatusMessage,
								i_etDiag		:= GD.ET_Diag.Ok,
								i_udiDiagExt	:= AXM_ET_DiagExt.Ok,
								i_sMessage		:= Standard.CONCAT(Standard.CONCAT(Standard.CONCAT('Command done: ', AXM_FC_EtCmdToString(i_etCmd := iq_stStandardModuleItf.iq_diCmd)),' number: '),DINT_TO_STRING(iq_stStandardModuleItf.iq_diCmd)),
								q_etDiag		:= ,
								q_etDiagExt		:= );
END_IF

iq_stStandardModuleItf.q_xCmdActive := FALSE;
iq_stStandardModuleItf.q_xCmdDone := TRUE;
IF(iq_stStandardModuleItf.iq_diCmd = iq_stStandardModuleItf.q_diCmdActive) THEN
	iq_stStandardModuleItf.iq_diCmd := 0;
(* ELSE don't touch iq_diCMD *)
END_IF

(* ---- SignalUnsuccessfulExecution.meth.st ---- *)
{attribute 'conditionalshow_all_locals'}
METHOD INTERNAL SignalUnsuccessfulExecution
VAR_INPUT
END_VAR

IF fbLoggerPoint.etLogLevel >= APL.ET_LogLevel.StatusMessage THEN
	fbLoggerPoint.AddLogEntry(	i_etLogLevel	:= APL.ET_LogLevel.StatusMessage,
								i_etDiag		:= GD.ET_Diag.Ok,
								i_udiDiagExt	:= AXM_ET_DiagExt.Ok,
								i_sMessage		:= Standard.CONCAT(Standard.CONCAT(Standard.CONCAT('Command failed: ', AXM_FC_EtCmdToString(i_etCmd := iq_stStandardModuleItf.iq_diCmd)),' number: '),DINT_TO_STRING(iq_stStandardModuleItf.iq_diCmd)),
								q_etDiag		:= ,
								q_etDiagExt		:= );
END_IF

iq_stStandardModuleItf.q_xCmdActive := FALSE;
iq_stStandardModuleItf.q_xCmdDone := FALSE;
IF(iq_stStandardModuleItf.iq_diCmd = iq_stStandardModuleItf.q_diCmdActive) THEN
	iq_stStandardModuleItf.iq_diCmd := -iq_stStandardModuleItf.iq_diCmd;
(* ELSE don't touch iq_diCMD *)
END_IF
